(*
SPDX-FileCopyrightText: c 2026 Oleksandr Tiutyk <trofimich@gmail.com>
SPDX-License-Identifier: MIT
License: https://opensource.org/license/mit
*)

(*!
<summary>Checks borrowed insertion and suffix order.</summary>
<description>
Borrows a group-owned list reserved for this case. Use from one task at a stable address.
Teardown clears the list before publication.
</description>
*)

{attribute 'no_assign'}
{attribute 'no_explicit_call' := 'do not call this function block directly'}
FUNCTION_BLOCK ListInsertGenericTest EXTENDS TOF_Testing.SingleCycleTest
VAR_STAT
	{attribute 'hide'}
	_ClassName : STRING := __POUNAME();
END_VAR
VAR
	_List : TOF_Collections.IList;
	_Values : ARRAY [0..5] OF STRING := ['String0', 'String1', 'String2', 'String3', 'String4', 'String5'];
END_VAR

(*!
<summary>Clears the fixture before the runner publishes the result.</summary>
<description>
Also runs after an unexpected exception interrupts the case.
</description>
*)
METHOD PROTECTED AfterTest
_List.Clear();
END_METHOD

//! <summary>Borrows the concrete class name. Callers must not modify it.</summary>
{attribute 'monitoring' := 'call'}
PROPERTY ClassName : REFERENCE TO STRING
GET
ClassName REF= _ClassName;
END_GET
END_PROPERTY

(*!
<summary>Checks borrowed insertion and suffix order.</summary>
*)
METHOD PROTECTED ExecuteTest
VAR
	values : ARRAY [0..5] OF STRING := ['String0', 'String1', 'String2', 'String3', 'String4', 'String5'];
	entry : TOF_Core.GENERIC_VALUE;
	expected : ARRAY [0..3] OF STRING := ['String0', 'String5', 'String1', 'String2'];
	i : DINT;
END_VAR
_List.AppendCopy(value := values[0]);
_List.AppendCopy(value := values[1]);
_List.AppendCopy(value := values[2]);

entry := TOF_Core.GenericValueFactory.FromStringReference(value := _Values[5]);
_List.InsertGeneric(index := 1, value := entry);

Assert.ThatBool(
	actual := _List.Get(index := 1).Address = entry.Address AND_THEN NOT _List.Get(index := 1).IsMemoryOwner,
	message := "InsertGeneric must retain the borrowed address and ownership mode"
).IsTrue();

Assert.ThatDInt(
	actual := _List.Length,
	message := "Unexpected sequence after InsertGeneric length"
).ToBe(expected := DINT#4);

FOR i := 0 TO 3 DO
	Assert.ThatString(
		actual := _List.Get(index := i).AsString255(),
		message := TOF_Core.WideStrings.Concat255("Unexpected sequence after InsertGeneric at index ", TO_WSTRING(i))
	).ToBe(expected := expected[i]);
END_FOR
END_METHOD

(*!
<summary>Binds the list fixture for this case.</summary>
<description>
Stores a borrowed interface without invoking the fixture. The owning group keeps it alive and
reserves it for this case. TestElement initializes the name and parent.
</description>
<param name="name">Display name of this case.</param>
<param name="parent">Group that owns this case.</param>
<param name="list">Required live list reserved for this case.</param>
*)
METHOD FB_init : BOOL
VAR_INPUT
	bInitRetains: BOOL; // TRUE: the retain variables are initialized (reset warm / reset cold)
	bInCopyCode: BOOL; // TRUE: the instance will be copied to the copy code afterward (online change)
	name : WSTRING;
	parent : TOF_Testing.ITestElement;
	list : TOF_Collections.IList;
END_VAR
_List := list;
FB_init := TRUE;
END_METHOD

//! <summary>Borrows the compiler-initialized namespace name. Callers must not modify it.</summary>
{attribute 'monitoring' := 'call'}
PROPERTY NamespaceName : REFERENCE TO STRING
GET
NamespaceName REF= CurrentNamespace.Name;
END_GET
END_PROPERTY

//! <summary>Reports the concrete instance size in bytes.</summary>
{attribute 'monitoring' := 'call'}
PROPERTY SelfSize : ULINT
GET
SelfSize := XSIZEOF(THIS^);
END_GET
END_PROPERTY

END_FUNCTION_BLOCK

(* stored: Version 1.1.0.1, ProductVersion 3.1.4026.21
   POU ListInsertGenericTest: Id {a891092b-b113-4fe5-b8df-2b790337f86c}, SpecialFunc None
   Method AfterTest: Id {d871ea64-d23b-4c82-aaeb-3d7dc9498a33}
   Property ClassName: Id {b9a445c9-0c26-41ea-83ef-4363970ae4f6}
   Get Get: Id {21f43e13-6a92-4502-8b5d-b0c4426fd9e8}
   Method ExecuteTest: Id {d98307c1-5348-4e4d-9f0f-b4026c96405b}
   Method FB_init: Id {57377cf7-f0ed-43b5-963c-952546b74892}
   Property NamespaceName: Id {ed790d17-072b-474b-9588-e7092f3bce22}
   Get Get: Id {93757623-7925-46bb-8a23-115ba1095b2d}
   Property SelfSize: Id {903528cb-512a-4514-bdea-aa43d59524ea}
   Get Get: Id {fe8e677f-5cc0-4a55-aace-251d18743d4d} *)
